(* IEC 61131-3 sources: crb-codesys/generation/scripts/repoeval/plc_hello_mixing_tank/struct, 2 files *)

(* ---- AUTO_SEQUENCE.st ---- *)
{attribute 'qualified_only' := ''}
{attribute 'strict' := ''}
TYPE AUTO_SEQUENCE :
(
	///Draining state when system is in auto mode
	DRAINING := 0,
	///Filling state when system is in auto mode
	FILLING := 1,
	///Mixing state when system is in auto mode
	MIXING := 2
);
END_TYPE

(* ---- MODES.st ---- *)
{attribute 'qualified_only' := ''}
{attribute 'strict' := ''}
TYPE MODES :
(
	///System is in manual mode (Operator control)
	MANUAL := 0,
	///System is in auto mode (PLC in control)
	AUTO := 1
);
END_TYPE
